FUNCTION_BLOCK FB_CoverControl IMPLEMENTS I_MirrorCovers
VAR_INPUT
	Delta		: TIME := T#5S;		// Time difference between both covers opening (and closing)
	TimeToCycle	: TIME := T#15S;	// Time for one motor to fully open/close
	// TRUE while the E-stop is triggered (MAIN: safetyHandling.estop): moving covers stop, open/close requests
	// are dropped (#15)
	bEmergency	: BOOL;
END_VAR
VAR_OUTPUT
END_VAR
VAR
	bOpen		: BOOL;
	bClose		: BOOL;
	bStop		: BOOL;
	// State
	fbCoverIdleState : FB_CoverIdleState(THIS);
	fbCoverOpeningState : FB_CoverOpeningState(THIS);
	fbCoverStoppingState : FB_CoverStoppingState(THIS);
	fbCoverClosingState : FB_CoverClosingState(THIS);
	
	ipState		: I_CoverState := fbCoverIdleState;
	// #111: the PLC cannot know the position of the covers after a start (activation, Reset Cold), so it starts with
	// "unknown" instead of assuming "closed". The first open or close cycle that completes sets the real end position.
	eCoverState	: E_MirrorCoverState := E_MirrorCoverState.unknown;
	// #71: TRUE only once an open or close cycle has completed since the PLC start. Until then the position is
	// unknown (the covers may be open after a restart), so a request is only ignored once the position is confirmed.
	bEndPositionConfirmed : BOOL := FALSE;
	bRequestIgnored : BOOL;
	// Trigger
	rtrigOpen		: R_TRIG;
	rtrigClose		: R_TRIG;
	rtrigStop		: R_TRIG;
	// Comm
	fbComm			: I_Comm;
	tonComm 		: TON := (PT:=T#5S);
	fbCoverOpenEvent:	FB_EventLog;
	fbCoverClosedEvent: FB_EventLog;
	fbCoverEmergencyEvent: FB_EventLog;
	fbCoverIgnoredEvent: FB_EventLog;
	// Motor relais
	bMotor1RelaisA	AT%Q*	: BOOL := FALSE;
	bMotor1RelaisB	AT%Q*	: BOOL := FALSE;
	
	bMotor2RelaisA	AT%Q*	: BOOL := FALSE;
	bMotor2RelaisB	AT%Q*	: BOOL := FALSE;
END_VAR

rtrigOpen(CLK := bOpen);
rtrigClose(CLK := bClose);
rtrigStop(CLK := bStop);
bRequestIgnored := FALSE;

IF bEmergency THEN
	// requests made during the E-stop are dropped (flags cleared below, #15)
	// stop only moving covers, so that closed/open covers keep their known state
	IF eCoverState = E_MirrorCoverState.opening OR eCoverState = E_MirrorCoverState.closing THEN
		ipState.StopCommand();
	END_IF
ELSE
	IF rtrigStop.Q THEN
		ipState.StopCommand();
	END_IF

	// #71: a request for the position the covers are confirmed to be in does nothing (it ran a full 20 s cycle)
	IF rtrigClose.Q THEN
		IF eCoverState = E_MirrorCoverState.closed AND bEndPositionConfirmed THEN
			bRequestIgnored := TRUE;
		ELSE
			ipState.CloseCommand();
		END_IF
	END_IF

	IF rtrigOpen.Q THEN
		IF eCoverState = E_MirrorCoverState.open AND bEndPositionConfirmed THEN
			bRequestIgnored := TRUE;
		ELSE
			ipState.OpenCommand();
		END_IF
	END_IF
END_IF

// #66: requests are one-shot. They are consumed in this scan whether they produced an edge or not, so a caller that
// repeats a request every scan (the park, stage 80) cannot leave a flag TRUE: left set, it would block the rising
// edge of every later request.
bOpen := FALSE;
bClose := FALSE;
bStop := FALSE;

ipState.RunState();

// send telemetry
tonComm(IN:=TRUE);
IF tonComm.Q THEN // publish new payload every second
	tonComm(IN:=FALSE);
	THIS^._SendTelemetry();	
END_IF


fbCoverOpenEvent(
	Trigger := eCoverState = E_MirrorCoverState.open,
	Level := ADSLOG_MSGTYPE_HINT,
	OnMessage := 'Mirror cover is open.',
	comm:= fbComm);
fbCoverClosedEvent(
	Trigger := eCoverState = E_MirrorCoverState.closed,
	Level := ADSLOG_MSGTYPE_HINT,
	OnMessage := 'Mirror cover is closed.',
	comm:= fbComm);
fbCoverIgnoredEvent(
	Trigger := bRequestIgnored,
	Level := ADSLOG_MSGTYPE_HINT,
	OnMessage := 'Mirror cover already in the requested end position, request ignored.',
	comm:= fbComm);
fbCoverEmergencyEvent(
	Trigger := bEmergency,
	Level := ADSLOG_MSGTYPE_WARN,
	OnMessage := 'Mirror cover: E-stop, covers stopped and commands ignored.',
	comm:= fbComm);

PROPERTY _CoverState : E_MirrorCoverState
SET
eCoverState := _CoverState;
bEndPositionConfirmed := (_CoverState = E_MirrorCoverState.closed OR _CoverState = E_MirrorCoverState.open);
END_SET
END_PROPERTY

PROPERTY _Motor1RelaisA : BOOL
SET
bMotor1RelaisA := _Motor1RelaisA;
END_SET
END_PROPERTY

PROPERTY _Motor1RelaisB : BOOL
SET
bMotor1RelaisB := _Motor1RelaisB;
END_SET
END_PROPERTY

PROPERTY _Motor2RelaisA : BOOL
SET
bMotor2RelaisA := _Motor2RelaisA;
END_SET
END_PROPERTY

PROPERTY _Motor2RelaisB : BOOL
SET
bMotor2RelaisB := _Motor2RelaisB;
END_SET
END_PROPERTY

METHOD _SendTelemetry : BOOL
VAR_INPUT
END_VAR
IF eCoverState = E_MirrorCoverState.closed THEN
	fbComm.PublishLREAL('telescope', 'dome', 'AUXILIARY.COVER.REALPOS', 0.0);
ELSIF eCoverState = E_MirrorCoverState.open THEN
	fbComm.PublishLREAL('telescope', 'dome', 'AUXILIARY.COVER.REALPOS', 1.0);
ELSE
	// moving, stopped or unknown (#111): not at an end position
	fbComm.PublishLREAL('telescope', 'dome', 'AUXILIARY.COVER.REALPOS', 0.5);
END_IF
END_METHOD

METHOD Close : BOOL
VAR_INPUT
END_VAR
bClose := TRUE;
END_METHOD

PROPERTY Closed : BOOL
GET
IF THIS^.CoverState = E_MirrorCoverState.closed THEN
	Closed := TRUE;
ELSE
	Closed := FALSE;
END_IF
END_GET
END_PROPERTY

PROPERTY CoverState : E_MirrorCoverState
GET
CoverState := eCoverState;
END_GET
END_PROPERTY

PROPERTY Error : BOOL
GET
Error := FALSE;
END_GET
END_PROPERTY

//FB_Init is always available implicitly and it is used primarily for initialization.
//The return value is not evaluated. For a specific influence, you can also declare the
//methods explicitly and provide additional code there with the standard initialization
//code. You can evaluate the return value.
METHOD FB_Init: BOOL
VAR_INPUT
    bInitRetains	: BOOL; // TRUE: the retain variables are initialized (reset warm / reset cold)
    bInCopyCode		: BOOL;  // TRUE: the instance will be copied to the copy code afterward (online change)
	comm			: I_Comm;
END_VAR
THIS^.fbComm 				:= comm;
END_METHOD

METHOD Open : BOOL
VAR_INPUT
END_VAR
bOpen := TRUE;
END_METHOD

PROPERTY Opened : BOOL
GET
IF THIS^.CoverState = E_MirrorCoverState.open THEN
	Opened := TRUE;
ELSE
	Opened := FALSE;
END_IF
END_GET
END_PROPERTY

METHOD Reset : BOOL
VAR_INPUT
END_VAR
END_METHOD

METHOD SetState : BOOL
VAR_INPUT
	newState :I_CoverState;
END_VAR
THIS^.ipState := newState;
END_METHOD

METHOD Stop : BOOL
VAR_INPUT
END_VAR
bStop := TRUE;
END_METHOD

END_FUNCTION_BLOCK

(* stored: Version 1.1.0.1, ProductVersion 3.1.4024.15
   POU FB_CoverControl: Id {d3621f5c-b414-4287-a5b0-c413b9f4d1e9}, SpecialFunc None
   Folder internal properties: Id {d7d68b3e-5318-439e-87f9-1ef435c0c5d1}
   Folder properties: Id {aaac3f27-dfda-472e-bc85-10fb56c84bfd}
   Property _CoverState: Id {c85b32fd-9415-4791-974c-4ca08103afd7}
   Set Set: Id {f51f43d2-3fdd-457e-81b4-6e2279702ecb}
   Property _Motor1RelaisA: Id {a8604255-4e83-4e3e-bb1b-8fa1f8af3270}
   Set Set: Id {f7b1a4d7-2ab8-4214-9701-469cce4c1746}
   Property _Motor1RelaisB: Id {c75eed28-e932-4804-a2fa-76dad7b24886}
   Set Set: Id {c28745b5-4222-499c-a64f-4847f3da5bd5}
   Property _Motor2RelaisA: Id {c44f1da8-f693-4b7b-9269-3c0e57eaede2}
   Set Set: Id {a5d54a7c-47dd-415c-bf54-8e1d77599bd1}
   Property _Motor2RelaisB: Id {b776bd98-83fd-4b81-b3ec-6d518283dd14}
   Set Set: Id {99aa748e-7bd2-4d38-9d81-f8812add68c4}
   Method _SendTelemetry: Id {0a8e627f-9fae-40e1-bd53-318ad436c233}
   Method Close: Id {0a475567-f0d9-4b8f-a207-512f31f9b819}
   Property Closed: Id {fe324a82-ce87-4c62-a8bf-44fbeb3a3228}
   Get Get: Id {7e2dccd8-daa7-43a8-bdab-75dce67348c4}
   Property CoverState: Id {9900c09a-8af5-4aa1-819a-8a64815ba24c}
   Get Get: Id {b1274ca8-7d60-4a57-b23e-6e172401778c}
   Property Error: Id {d53107c8-e453-4e05-bc9a-229014b7917d}
   Get Get: Id {a72e4b0a-3a23-4243-9719-6e644c76db05}
   Method FB_Init: Id {29f2f728-7391-4fd0-b6a5-8535dccce95b}
   Method Open: Id {ab86d33d-a775-4eaa-8b2e-bcc3ba9a3c80}
   Property Opened: Id {5f095883-e244-4fba-b20f-8b0ae1386b52}
   Get Get: Id {3e705fa8-212a-4465-a041-b00481831e3c}
   Method Reset: Id {ab37cc4b-70b9-4d04-96df-5f7175bb7ce3}
   Method SetState: Id {1dc7bcb9-616a-44a2-977b-f8fb97eb2447}
   Method Stop: Id {a261d6e5-60ee-4a27-9286-882b77ec4095} *)
